// TIA Portal V20 export
// export: Created 2026-10-20T12:51:00.7155082Z, ExportSetting WithDefaults, DisplayName Totally Integrated Automation Portal, DisplayVersion V20 Update 6, DisplayName TIA Portal Openness, DisplayVersion V20 Update 6, DisplayName TIA Portal Version Control Interface, DisplayVersion V20 Update 6, DisplayName SINAMICS Startdrive Advanced, DisplayVersion V20 SP1, DisplayName SINAMICS Startdrive G130, G150, S120, S150, SINAMICS MV, G220, S200, S210, DisplayVersion V20 SP1, DisplayName SINAMICS Startdrive G110M, G120, G120C, G120D, G120P, G115D, DisplayVersion V20 SP1, DisplayName STEP 7 Professional, DisplayVersion V20 Update 6, DisplayName STEP 7 Safety, DisplayVersion V20 Update 2, DisplayName WinCC Basic/Comfort/Advanced, DisplayVersion V20 Update 6, DisplayName WinCC Unified, DisplayVersion V20 Update 6
FUNCTION_BLOCK "F_Lock_FB"   // FB24, F_FBD
{ S7_Optimized_Access := 'TRUE' }
VERSION : 0.1
// stored: AutoNumber true, IsIECCheckEnabled false, UDAEnableTagReadback false
   VAR_INPUT
      Lock_Closed_CH1 { ExternalAccessible := 'False'; ExternalVisible := 'False'; ExternalWritable := 'False'} : Bool;
      Lock_Closed_CH2 { ExternalAccessible := 'False'; ExternalVisible := 'False'; ExternalWritable := 'False'} : Bool;
      EStop_CH1 { ExternalAccessible := 'False'; ExternalVisible := 'False'; ExternalWritable := 'False'} : Bool;
      EStop_CH2 { ExternalAccessible := 'False'; ExternalVisible := 'False'; ExternalWritable := 'False'} : Bool;
      ACK { ExternalAccessible := 'False'; ExternalVisible := 'False'; ExternalWritable := 'False'} : Bool;
   END_VAR
   VAR_OUTPUT
      Lock_Reset_Input1 { ExternalAccessible := 'False'; ExternalVisible := 'False'; ExternalWritable := 'False'} : Bool;
      Lock_Reset_Input2 { ExternalAccessible := 'False'; ExternalVisible := 'False'; ExternalWritable := 'False'} : Bool;
      Lock_Reset_Input3 { ExternalAccessible := 'False'; ExternalVisible := 'False'; ExternalWritable := 'False'} : Bool;
      Lock_Reset_Input4 { ExternalAccessible := 'False'; ExternalVisible := 'False'; ExternalWritable := 'False'} : Bool;
      EStop_Lock_OK : Bool;
      Lock_Secured_OK : Bool;
   END_VAR
   VAR
      GUARD_SWITCH : ESTOP1;
      ESTOP : ESTOP1;
   END_VAR
BEGIN

REGION Network 1: GUARD SWITCH
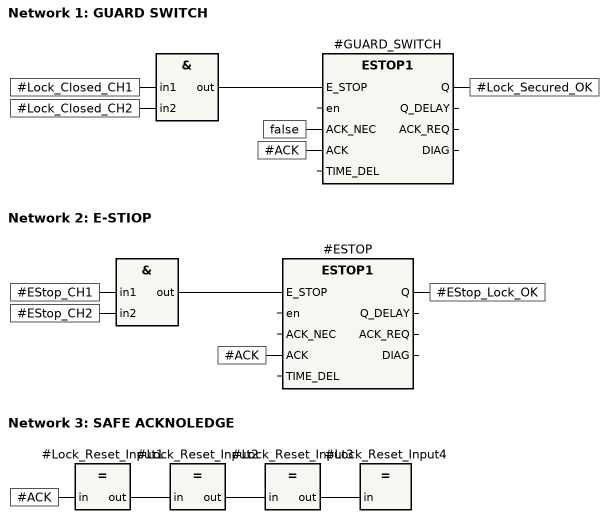
   #GUARD_SWITCH(E_STOP := #Lock_Closed_CH1 AND #Lock_Closed_CH2,   // ESTOP1
                 ACK_NEC := false,
                 ACK := #ACK,
                 Q => #Lock_Secured_OK);
END_REGION

REGION Network 2: E-STIOP
   #ESTOP(E_STOP := #EStop_CH1 AND #EStop_CH2, ACK := #ACK, Q => #EStop_Lock_OK);   // ESTOP1
END_REGION

REGION Network 3: SAFE ACKNOLEDGE
   #Lock_Reset_Input1 := #ACK;
   #Lock_Reset_Input2 := #ACK;
   #Lock_Reset_Input3 := #ACK;
   #Lock_Reset_Input4 := #ACK;
END_REGION
END_FUNCTION_BLOCK
